(* IEC 61131-3 sources: plc-workbench/examples/motor/mutants, 3 files *)

(* ---- ignore_estop.st ---- *)
(* SYNTHETIC FAULT: ignore_estop -- deliberately incorrect. *)
FUNCTION_BLOCK MotorControl
VAR_INPUT
    StartBtn : BOOL;
    StopBtn : BOOL;
    EStop : BOOL;
END_VAR
VAR_OUTPUT
    Motor : BOOL := FALSE;
END_VAR
IF StopBtn THEN
    Motor := FALSE;
ELSIF StartBtn THEN
    Motor := TRUE;
END_IF;
END_FUNCTION_BLOCK

(* ---- lost_latch.st ---- *)
(* SYNTHETIC FAULT: lost_latch -- deliberately incorrect. *)
FUNCTION_BLOCK MotorControl
VAR_INPUT
    StartBtn : BOOL;
    StopBtn : BOOL;
    EStop : BOOL;
END_VAR
VAR_OUTPUT
    Motor : BOOL := FALSE;
END_VAR
IF StopBtn OR EStop THEN
    Motor := FALSE;
ELSIF StartBtn THEN
    Motor := TRUE;
ELSE
    Motor := FALSE;
END_IF;
END_FUNCTION_BLOCK

(* ---- start_over_stop.st ---- *)
(* SYNTHETIC FAULT: start_over_stop -- deliberately incorrect. *)
FUNCTION_BLOCK MotorControl
VAR_INPUT
    StartBtn : BOOL;
    StopBtn : BOOL;
    EStop : BOOL;
END_VAR
VAR_OUTPUT
    Motor : BOOL := FALSE;
END_VAR
IF StartBtn THEN
    Motor := TRUE;
ELSIF StopBtn OR EStop THEN
    Motor := FALSE;
END_IF;
END_FUNCTION_BLOCK
